FUNCTION_BLOCK RoboCat (* CAT Function Block Type *)
  (* Standard: 61499-2 *)
  (* Version 0.0, 7/10/2026, template *)
  PACKAGE Main;
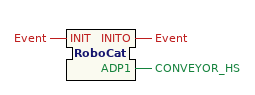
  EVENT_INPUT
    INIT; (* Initialization Request *)
  END_EVENT
  EVENT_OUTPUT
    INITO; (* Initialization Confirm *)
  END_EVENT
  PLUGS
    ADP1 : CONVEYOR_HS;
  END_PLUGS
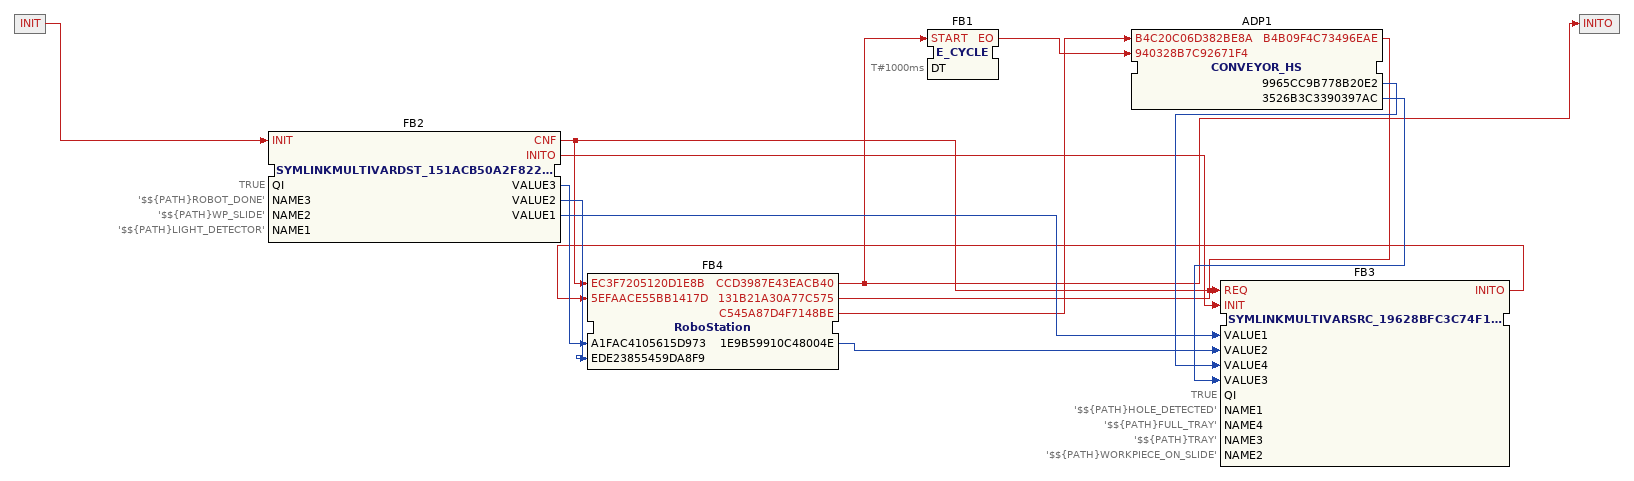
  FBS
    FB1 : E_CYCLE(DT := T#1000ms);
    FB2 : SYMLINKMULTIVARDST_151ACB50A2F8223B2(QI := TRUE, NAME3 := '$${PATH}ROBOT_DONE', NAME2 := '$${PATH}WP_SLIDE', NAME1 := '$${PATH}LIGHT_DETECTOR'); {SET_ATTRIBUTE(Configuration.GenericFBType.InterfaceParams, Runtime.System#I:=3;VALUE${I$}:BOOL,BOOL,BOOL)}
    FB3 : SYMLINKMULTIVARSRC_19628BFC3C74F1AB1(QI := TRUE, NAME1 := '$${PATH}HOLE_DETECTED', NAME4 := '$${PATH}FULL_TRAY', NAME3 := '$${PATH}TRAY', NAME2 := '$${PATH}WORKPIECE_ON_SLIDE'); {SET_ATTRIBUTE(Configuration.GenericFBType.InterfaceParams, Runtime.System#I:=4;VALUE${I$}:BOOL,BOOL,BOOL,BOOL)}
    FB4 : RoboStation;
  END_FBS
  EVENT_CONNECTIONS
    INIT TO FB2.INIT;
    FB2.CNF TO FB4.EC3F7205120D1E8B;
    FB2.CNF TO FB3.REQ;
    ADP1.B4B09F4C73496EAE TO FB3.REQ;
    FB2.INITO TO FB3.INIT;
    FB3.INITO TO FB4.5EFAACE55BB1417D;
    FB4.CCD3987E43EACB40 TO FB1.START;
    FB4.CCD3987E43EACB40 TO INITO;
    FB4.131B21A30A77C575 TO FB3.REQ;
    FB4.C545A87D4F7148BE TO ADP1.B4C20C06D382BE8A;
    FB1.EO TO ADP1.940328B7C92671F4;
  END_CONNECTIONS
  DATA_CONNECTIONS
    FB2.VALUE3 TO FB4.A1FAC4105615D973;
    FB2.VALUE2 TO FB4.EDE23855459DA8F9;
    FB2.VALUE1 TO FB3.VALUE1;
    FB4.1E9B59910C48004E TO FB3.VALUE2;
    ADP1.9965CC9B778B20E2 TO FB3.VALUE4;
    ADP1.3526B3C3390397AC TO FB3.VALUE3;
  END_CONNECTIONS
END_FUNCTION_BLOCK
